Omron CX-Programmer project NewProject (CX-Programmer 9.51)

# PLC NewPLC1: CP1L L

## Global symbols (name address type ; comment)
W0.01 BOOL  ; \

## Program NewProgram1 (cyclic task 0)
Local symbols
button_1 0.00 BOOL
button_2 0.02 BOOL
button_3 0.04 BOOL
out_1 100.00 BOOL
out_2 100.01 BOOL
out_3 100.02 BOOL

### Section Section1

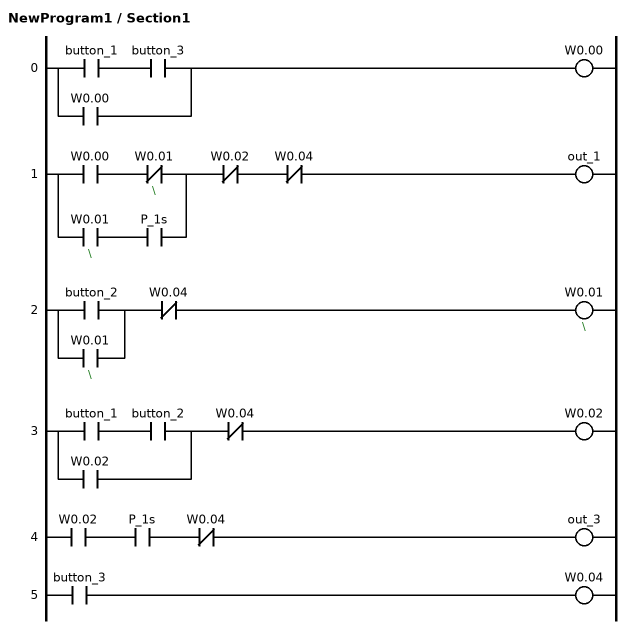
; rung 0
LD button_1
AND button_3
OR W0.00
OUT W0.00
; rung 1
LD W0.00
ANDNOT W0.01  ; \
LD W0.01  ; \
AND P_1s
ORLD
ANDNOT W0.02
ANDNOT W0.04
OUT out_1
; rung 2
LD button_2
OR W0.01  ; \
ANDNOT W0.04
OUT W0.01  ; \
; rung 3
LD button_1
AND button_2
OR W0.02
ANDNOT W0.04
OUT W0.02
; rung 4
LD W0.02
AND P_1s
ANDNOT W0.04
OUT out_3
; rung 5
LD button_3
OUT W0.04

### Section END
; rung 0
END(001)